FUNCTION "FRK_PersistRootStatus" : Void
{ S7_Optimized_Access := 'TRUE' }
VERSION : 0.1
VAR_INPUT
    RootIndex : Int;
END_VAR
VAR_IN_OUT
    Persist : "ST_ConfigPersistStatus";
END_VAR
BEGIN
    IF #RootIndex < 1 OR #RootIndex > 2 THEN RETURN; END_IF;
    #Persist.Pending := FALSE; #Persist.PendingSince := LDT#1970-01-01-00:00:00;
    #Persist.WindowMs := 26000;
    IF #RootIndex = 1 THEN
        #Persist.Failed := #Persist.Failed OR "FRK_PersistConsumers".Rows[1].Failed;
        IF "FRK_PersistConsumers".Rows[1].Dirty OR "FRK_PersistConsumers".Rows[1].Ticket <> 0 THEN
            #Persist.Pending := TRUE;
            IF #Persist.PendingSince = LDT#1970-01-01-00:00:00 OR ("FRK_PersistConsumers".Rows[1].PendingSince <> LDT#1970-01-01-00:00:00 AND "FRK_PersistConsumers".Rows[1].PendingSince < #Persist.PendingSince) THEN #Persist.PendingSince := "FRK_PersistConsumers".Rows[1].PendingSince; END_IF;
        END_IF;
    END_IF;
    IF #RootIndex = 1 THEN
        #Persist.Failed := #Persist.Failed OR "FRK_PersistConsumers".Rows[2].Failed;
        IF "FRK_PersistConsumers".Rows[2].Dirty OR "FRK_PersistConsumers".Rows[2].Ticket <> 0 THEN
            #Persist.Pending := TRUE;
            IF #Persist.PendingSince = LDT#1970-01-01-00:00:00 OR ("FRK_PersistConsumers".Rows[2].PendingSince <> LDT#1970-01-01-00:00:00 AND "FRK_PersistConsumers".Rows[2].PendingSince < #Persist.PendingSince) THEN #Persist.PendingSince := "FRK_PersistConsumers".Rows[2].PendingSince; END_IF;
        END_IF;
    END_IF;
    IF #RootIndex = 1 THEN
        #Persist.Failed := #Persist.Failed OR "FRK_PersistConsumers".Rows[3].Failed;
        IF "FRK_PersistConsumers".Rows[3].Dirty OR "FRK_PersistConsumers".Rows[3].Ticket <> 0 THEN
            #Persist.Pending := TRUE;
            IF #Persist.PendingSince = LDT#1970-01-01-00:00:00 OR ("FRK_PersistConsumers".Rows[3].PendingSince <> LDT#1970-01-01-00:00:00 AND "FRK_PersistConsumers".Rows[3].PendingSince < #Persist.PendingSince) THEN #Persist.PendingSince := "FRK_PersistConsumers".Rows[3].PendingSince; END_IF;
        END_IF;
    END_IF;
    IF #RootIndex = 1 THEN
        #Persist.Failed := #Persist.Failed OR "FRK_PersistConsumers".Rows[4].Failed;
        IF "FRK_PersistConsumers".Rows[4].Dirty OR "FRK_PersistConsumers".Rows[4].Ticket <> 0 THEN
            #Persist.Pending := TRUE;
            IF #Persist.PendingSince = LDT#1970-01-01-00:00:00 OR ("FRK_PersistConsumers".Rows[4].PendingSince <> LDT#1970-01-01-00:00:00 AND "FRK_PersistConsumers".Rows[4].PendingSince < #Persist.PendingSince) THEN #Persist.PendingSince := "FRK_PersistConsumers".Rows[4].PendingSince; END_IF;
        END_IF;
    END_IF;
    IF #RootIndex = 1 THEN
        #Persist.Failed := #Persist.Failed OR "FRK_PersistConsumers".Rows[5].Failed;
        IF "FRK_PersistConsumers".Rows[5].Dirty OR "FRK_PersistConsumers".Rows[5].Ticket <> 0 THEN
            #Persist.Pending := TRUE;
            IF #Persist.PendingSince = LDT#1970-01-01-00:00:00 OR ("FRK_PersistConsumers".Rows[5].PendingSince <> LDT#1970-01-01-00:00:00 AND "FRK_PersistConsumers".Rows[5].PendingSince < #Persist.PendingSince) THEN #Persist.PendingSince := "FRK_PersistConsumers".Rows[5].PendingSince; END_IF;
        END_IF;
    END_IF;
    IF #RootIndex = 1 THEN
        #Persist.Failed := #Persist.Failed OR "FRK_PersistConsumers".Rows[6].Failed;
        IF "FRK_PersistConsumers".Rows[6].Dirty OR "FRK_PersistConsumers".Rows[6].Ticket <> 0 THEN
            #Persist.Pending := TRUE;
            IF #Persist.PendingSince = LDT#1970-01-01-00:00:00 OR ("FRK_PersistConsumers".Rows[6].PendingSince <> LDT#1970-01-01-00:00:00 AND "FRK_PersistConsumers".Rows[6].PendingSince < #Persist.PendingSince) THEN #Persist.PendingSince := "FRK_PersistConsumers".Rows[6].PendingSince; END_IF;
        END_IF;
    END_IF;
    IF #RootIndex = 1 THEN
        #Persist.Failed := #Persist.Failed OR "FRK_PersistConsumers".Rows[7].Failed;
        IF "FRK_PersistConsumers".Rows[7].Dirty OR "FRK_PersistConsumers".Rows[7].Ticket <> 0 THEN
            #Persist.Pending := TRUE;
            IF #Persist.PendingSince = LDT#1970-01-01-00:00:00 OR ("FRK_PersistConsumers".Rows[7].PendingSince <> LDT#1970-01-01-00:00:00 AND "FRK_PersistConsumers".Rows[7].PendingSince < #Persist.PendingSince) THEN #Persist.PendingSince := "FRK_PersistConsumers".Rows[7].PendingSince; END_IF;
        END_IF;
    END_IF;
    IF #RootIndex = 1 THEN
        #Persist.Failed := #Persist.Failed OR "FRK_PersistConsumers".Rows[8].Failed;
        IF "FRK_PersistConsumers".Rows[8].Dirty OR "FRK_PersistConsumers".Rows[8].Ticket <> 0 THEN
            #Persist.Pending := TRUE;
            IF #Persist.PendingSince = LDT#1970-01-01-00:00:00 OR ("FRK_PersistConsumers".Rows[8].PendingSince <> LDT#1970-01-01-00:00:00 AND "FRK_PersistConsumers".Rows[8].PendingSince < #Persist.PendingSince) THEN #Persist.PendingSince := "FRK_PersistConsumers".Rows[8].PendingSince; END_IF;
        END_IF;
    END_IF;
    IF #RootIndex = 2 THEN
        #Persist.Failed := #Persist.Failed OR "FRK_PersistConsumers".Rows[9].Failed;
        IF "FRK_PersistConsumers".Rows[9].Dirty OR "FRK_PersistConsumers".Rows[9].Ticket <> 0 THEN
            #Persist.Pending := TRUE;
            IF #Persist.PendingSince = LDT#1970-01-01-00:00:00 OR ("FRK_PersistConsumers".Rows[9].PendingSince <> LDT#1970-01-01-00:00:00 AND "FRK_PersistConsumers".Rows[9].PendingSince < #Persist.PendingSince) THEN #Persist.PendingSince := "FRK_PersistConsumers".Rows[9].PendingSince; END_IF;
        END_IF;
    END_IF;
    IF #RootIndex = 2 THEN
        #Persist.Failed := #Persist.Failed OR "FRK_PersistConsumers".Rows[10].Failed;
        IF "FRK_PersistConsumers".Rows[10].Dirty OR "FRK_PersistConsumers".Rows[10].Ticket <> 0 THEN
            #Persist.Pending := TRUE;
            IF #Persist.PendingSince = LDT#1970-01-01-00:00:00 OR ("FRK_PersistConsumers".Rows[10].PendingSince <> LDT#1970-01-01-00:00:00 AND "FRK_PersistConsumers".Rows[10].PendingSince < #Persist.PendingSince) THEN #Persist.PendingSince := "FRK_PersistConsumers".Rows[10].PendingSince; END_IF;
        END_IF;
    END_IF;
    IF #RootIndex = 2 THEN
        #Persist.Failed := #Persist.Failed OR "FRK_PersistConsumers".Rows[11].Failed;
        IF "FRK_PersistConsumers".Rows[11].Dirty OR "FRK_PersistConsumers".Rows[11].Ticket <> 0 THEN
            #Persist.Pending := TRUE;
            IF #Persist.PendingSince = LDT#1970-01-01-00:00:00 OR ("FRK_PersistConsumers".Rows[11].PendingSince <> LDT#1970-01-01-00:00:00 AND "FRK_PersistConsumers".Rows[11].PendingSince < #Persist.PendingSince) THEN #Persist.PendingSince := "FRK_PersistConsumers".Rows[11].PendingSince; END_IF;
        END_IF;
    END_IF;
    IF #RootIndex = 2 THEN
        #Persist.Failed := #Persist.Failed OR "FRK_PersistConsumers".Rows[12].Failed;
        IF "FRK_PersistConsumers".Rows[12].Dirty OR "FRK_PersistConsumers".Rows[12].Ticket <> 0 THEN
            #Persist.Pending := TRUE;
            IF #Persist.PendingSince = LDT#1970-01-01-00:00:00 OR ("FRK_PersistConsumers".Rows[12].PendingSince <> LDT#1970-01-01-00:00:00 AND "FRK_PersistConsumers".Rows[12].PendingSince < #Persist.PendingSince) THEN #Persist.PendingSince := "FRK_PersistConsumers".Rows[12].PendingSince; END_IF;
        END_IF;
    END_IF;
    IF #RootIndex = 2 THEN
        #Persist.Failed := #Persist.Failed OR "FRK_PersistConsumers".Rows[13].Failed;
        IF "FRK_PersistConsumers".Rows[13].Dirty OR "FRK_PersistConsumers".Rows[13].Ticket <> 0 THEN
            #Persist.Pending := TRUE;
            IF #Persist.PendingSince = LDT#1970-01-01-00:00:00 OR ("FRK_PersistConsumers".Rows[13].PendingSince <> LDT#1970-01-01-00:00:00 AND "FRK_PersistConsumers".Rows[13].PendingSince < #Persist.PendingSince) THEN #Persist.PendingSince := "FRK_PersistConsumers".Rows[13].PendingSince; END_IF;
        END_IF;
    END_IF;
    IF #RootIndex = 2 THEN
        #Persist.Failed := #Persist.Failed OR "FRK_PersistConsumers".Rows[14].Failed;
        IF "FRK_PersistConsumers".Rows[14].Dirty OR "FRK_PersistConsumers".Rows[14].Ticket <> 0 THEN
            #Persist.Pending := TRUE;
            IF #Persist.PendingSince = LDT#1970-01-01-00:00:00 OR ("FRK_PersistConsumers".Rows[14].PendingSince <> LDT#1970-01-01-00:00:00 AND "FRK_PersistConsumers".Rows[14].PendingSince < #Persist.PendingSince) THEN #Persist.PendingSince := "FRK_PersistConsumers".Rows[14].PendingSince; END_IF;
        END_IF;
    END_IF;
    IF #RootIndex = 2 THEN
        #Persist.Failed := #Persist.Failed OR "FRK_PersistConsumers".Rows[15].Failed;
        IF "FRK_PersistConsumers".Rows[15].Dirty OR "FRK_PersistConsumers".Rows[15].Ticket <> 0 THEN
            #Persist.Pending := TRUE;
            IF #Persist.PendingSince = LDT#1970-01-01-00:00:00 OR ("FRK_PersistConsumers".Rows[15].PendingSince <> LDT#1970-01-01-00:00:00 AND "FRK_PersistConsumers".Rows[15].PendingSince < #Persist.PendingSince) THEN #Persist.PendingSince := "FRK_PersistConsumers".Rows[15].PendingSince; END_IF;
        END_IF;
    END_IF;
    IF #RootIndex = 2 THEN
        #Persist.Failed := #Persist.Failed OR "FRK_PersistConsumers".Rows[16].Failed;
        IF "FRK_PersistConsumers".Rows[16].Dirty OR "FRK_PersistConsumers".Rows[16].Ticket <> 0 THEN
            #Persist.Pending := TRUE;
            IF #Persist.PendingSince = LDT#1970-01-01-00:00:00 OR ("FRK_PersistConsumers".Rows[16].PendingSince <> LDT#1970-01-01-00:00:00 AND "FRK_PersistConsumers".Rows[16].PendingSince < #Persist.PendingSince) THEN #Persist.PendingSince := "FRK_PersistConsumers".Rows[16].PendingSince; END_IF;
        END_IF;
    END_IF;

        #Persist.Failed := #Persist.Failed OR "FRK_PersistConsumers".Rows[17].Failed;
        IF "FRK_PersistConsumers".Rows[17].Dirty OR "FRK_PersistConsumers".Rows[17].Ticket <> 0 THEN
            #Persist.Pending := TRUE;
            IF #Persist.PendingSince = LDT#1970-01-01-00:00:00 OR ("FRK_PersistConsumers".Rows[17].PendingSince <> LDT#1970-01-01-00:00:00 AND "FRK_PersistConsumers".Rows[17].PendingSince < #Persist.PendingSince) THEN #Persist.PendingSince := "FRK_PersistConsumers".Rows[17].PendingSince; END_IF;
        END_IF;
    IF #RootIndex = 1 OR #RootIndex = 2 THEN
        #Persist.Failed := #Persist.Failed OR "FRK_PersistConsumers".Rows[18].Failed;
        IF "FRK_PersistConsumers".Rows[18].Dirty OR "FRK_PersistConsumers".Rows[18].Ticket <> 0 THEN
            #Persist.Pending := TRUE;
            IF #Persist.PendingSince = LDT#1970-01-01-00:00:00 OR ("FRK_PersistConsumers".Rows[18].PendingSince <> LDT#1970-01-01-00:00:00 AND "FRK_PersistConsumers".Rows[18].PendingSince < #Persist.PendingSince) THEN #Persist.PendingSince := "FRK_PersistConsumers".Rows[18].PendingSince; END_IF;
        END_IF;
    END_IF;
    IF (#RootIndex = 1 OR #RootIndex = 2) AND "FRK_PersistConsumers".Rows[18].Rejected AND NOT "FRK_PersistConsumers".Rows[18].Acknowledged THEN
        #Persist.RestoreLost := TRUE; #Persist.RestoreAcknowledged := FALSE;
        #Persist.LostPath := 'BenchLineOwner';
    END_IF;
    IF #RootIndex = 1 THEN
        #Persist.Failed := #Persist.Failed OR "FRK_PersistConsumers".Rows[19].Failed;
        IF "FRK_PersistConsumers".Rows[19].Dirty OR "FRK_PersistConsumers".Rows[19].Ticket <> 0 THEN
            #Persist.Pending := TRUE;
            IF #Persist.PendingSince = LDT#1970-01-01-00:00:00 OR ("FRK_PersistConsumers".Rows[19].PendingSince <> LDT#1970-01-01-00:00:00 AND "FRK_PersistConsumers".Rows[19].PendingSince < #Persist.PendingSince) THEN #Persist.PendingSince := "FRK_PersistConsumers".Rows[19].PendingSince; END_IF;
        END_IF;
    END_IF;
    IF #RootIndex = 2 THEN
        #Persist.Failed := #Persist.Failed OR "FRK_PersistConsumers".Rows[20].Failed;
        IF "FRK_PersistConsumers".Rows[20].Dirty OR "FRK_PersistConsumers".Rows[20].Ticket <> 0 THEN
            #Persist.Pending := TRUE;
            IF #Persist.PendingSince = LDT#1970-01-01-00:00:00 OR ("FRK_PersistConsumers".Rows[20].PendingSince <> LDT#1970-01-01-00:00:00 AND "FRK_PersistConsumers".Rows[20].PendingSince < #Persist.PendingSince) THEN #Persist.PendingSince := "FRK_PersistConsumers".Rows[20].PendingSince; END_IF;
        END_IF;
    END_IF;
    IF #Persist.Pending THEN
        IF "FRK_PersistRootSince".WasPending[#RootIndex] THEN
            IF "FRK_Elapsed"(NewMs := "FRK_Clock".NowMs, OldMs := "FRK_PersistRootSince".SinceMs[#RootIndex]) > #Persist.WindowMs THEN #Persist.Failed := TRUE; END_IF;
        ELSE "FRK_PersistRootSince".SinceMs[#RootIndex] := "FRK_Clock".NowMs; END_IF;
    END_IF;
    "FRK_PersistRootSince".WasPending[#RootIndex] := #Persist.Pending;
END_FUNCTION
FUNCTION "FRK_PersistAckRoot" : Void
{ S7_Optimized_Access := 'TRUE' }
VERSION : 0.1
VAR_INPUT
    RootIndex : Int;
END_VAR
BEGIN
    IF #RootIndex = 1 AND "FRK_PersistConsumers".Rows[1].Rejected THEN
        "FRK_PersistConsumers".Rows[1].Acknowledged := TRUE;
        "FRK_PersistRepair"(Slot := 1);
        "FRK_PersistDirty"(Slot := 1);
    END_IF;
    IF #RootIndex = 1 AND "FRK_PersistConsumers".Rows[2].Rejected THEN
        "FRK_PersistConsumers".Rows[2].Acknowledged := TRUE;
        "FRK_PersistRepair"(Slot := 2);
        "FRK_PersistDirty"(Slot := 2);
    END_IF;
    IF #RootIndex = 1 AND "FRK_PersistConsumers".Rows[3].Rejected THEN
        "FRK_PersistConsumers".Rows[3].Acknowledged := TRUE;
        "FRK_PersistRepair"(Slot := 3);
        "FRK_PersistDirty"(Slot := 3);
    END_IF;
    IF #RootIndex = 1 AND "FRK_PersistConsumers".Rows[4].Rejected THEN
        "FRK_PersistConsumers".Rows[4].Acknowledged := TRUE;
        "FRK_PersistRepair"(Slot := 4);
        "FRK_PersistDirty"(Slot := 4);
    END_IF;
    IF #RootIndex = 1 AND "FRK_PersistConsumers".Rows[5].Rejected THEN
        "FRK_PersistConsumers".Rows[5].Acknowledged := TRUE;
        "FRK_PersistRepair"(Slot := 5);
        "FRK_PersistDirty"(Slot := 5);
    END_IF;
    IF #RootIndex = 1 AND "FRK_PersistConsumers".Rows[6].Rejected THEN
        "FRK_PersistConsumers".Rows[6].Acknowledged := TRUE;
        "FRK_PersistRepair"(Slot := 6);
        "FRK_PersistDirty"(Slot := 6);
    END_IF;
    IF #RootIndex = 1 AND "FRK_PersistConsumers".Rows[7].Rejected THEN
        "FRK_PersistConsumers".Rows[7].Acknowledged := TRUE;
        "FRK_PersistRepair"(Slot := 7);
        "FRK_PersistDirty"(Slot := 7);
    END_IF;
    IF #RootIndex = 1 AND "FRK_PersistConsumers".Rows[8].Rejected THEN
        "FRK_PersistConsumers".Rows[8].Acknowledged := TRUE;
        "FRK_PersistRepair"(Slot := 8);
        "FRK_PersistDirty"(Slot := 8);
    END_IF;
    IF #RootIndex = 2 AND "FRK_PersistConsumers".Rows[9].Rejected THEN
        "FRK_PersistConsumers".Rows[9].Acknowledged := TRUE;
        "FRK_PersistRepair"(Slot := 9);
        "FRK_PersistDirty"(Slot := 9);
    END_IF;
    IF #RootIndex = 2 AND "FRK_PersistConsumers".Rows[10].Rejected THEN
        "FRK_PersistConsumers".Rows[10].Acknowledged := TRUE;
        "FRK_PersistRepair"(Slot := 10);
        "FRK_PersistDirty"(Slot := 10);
    END_IF;
    IF #RootIndex = 2 AND "FRK_PersistConsumers".Rows[11].Rejected THEN
        "FRK_PersistConsumers".Rows[11].Acknowledged := TRUE;
        "FRK_PersistRepair"(Slot := 11);
        "FRK_PersistDirty"(Slot := 11);
    END_IF;
    IF #RootIndex = 2 AND "FRK_PersistConsumers".Rows[12].Rejected THEN
        "FRK_PersistConsumers".Rows[12].Acknowledged := TRUE;
        "FRK_PersistRepair"(Slot := 12);
        "FRK_PersistDirty"(Slot := 12);
    END_IF;
    IF #RootIndex = 2 AND "FRK_PersistConsumers".Rows[13].Rejected THEN
        "FRK_PersistConsumers".Rows[13].Acknowledged := TRUE;
        "FRK_PersistRepair"(Slot := 13);
        "FRK_PersistDirty"(Slot := 13);
    END_IF;
    IF #RootIndex = 2 AND "FRK_PersistConsumers".Rows[14].Rejected THEN
        "FRK_PersistConsumers".Rows[14].Acknowledged := TRUE;
        "FRK_PersistRepair"(Slot := 14);
        "FRK_PersistDirty"(Slot := 14);
    END_IF;
    IF #RootIndex = 2 AND "FRK_PersistConsumers".Rows[15].Rejected THEN
        "FRK_PersistConsumers".Rows[15].Acknowledged := TRUE;
        "FRK_PersistRepair"(Slot := 15);
        "FRK_PersistDirty"(Slot := 15);
    END_IF;
    IF #RootIndex = 2 AND "FRK_PersistConsumers".Rows[16].Rejected THEN
        "FRK_PersistConsumers".Rows[16].Acknowledged := TRUE;
        "FRK_PersistRepair"(Slot := 16);
        "FRK_PersistDirty"(Slot := 16);
    END_IF;
    IF (#RootIndex = 1 OR #RootIndex = 2) AND "FRK_PersistConsumers".Rows[18].Rejected THEN
        "FRK_PersistConsumers".Rows[18].Acknowledged := TRUE;
        "FRK_PersistRepair"(Slot := 18);
        "FRK_PersistDirty"(Slot := 18);
    END_IF;
    IF (#RootIndex = 1 OR #RootIndex = 2) AND "FRK_PersistConsumers".Rows[18].Acknowledged AND "FRK_ConfigStore".LostPath[1] = 'BenchLineOwner' THEN
        "FRK_ConfigStore".Acknowledged[1] := TRUE;
    END_IF;
    IF #RootIndex = 1 AND "FRK_PersistConsumers".Rows[19].Rejected THEN
        "FRK_PersistConsumers".Rows[19].Acknowledged := TRUE;
        "FRK_PersistRepair"(Slot := 19);
        "FRK_PersistDirty"(Slot := 19);
    END_IF;
    IF #RootIndex = 2 AND "FRK_PersistConsumers".Rows[20].Rejected THEN
        "FRK_PersistConsumers".Rows[20].Acknowledged := TRUE;
        "FRK_PersistRepair"(Slot := 20);
        "FRK_PersistDirty"(Slot := 20);
    END_IF;
END_FUNCTION
